Fanuc KAREL source: KO00101.KL

PROGRAM KO00101
%NOLOCKGROUP
VAR
  A: INTEGER
  B: ARRAY[2] OF BYTE
  OUT: INTEGER
BEGIN
  A = 1
  B[1] = 2
  OUT = ATAN2(A, B[1])
END KO00101
